(* PLC project PR_ModeManageNoMode_PLC, SiemensToBackhoff Siemens TIA Portal to Beckhoff TwinCAT PLCopen Converter 1.0 *)
(* stored: creationDateTime 2026-09-28T08:41:48.575973Z, modificationDateTime 2026-09-28T08:41:48.575973Z *)

FUNCTION_BLOCK PR_ModeManageNoMode

(* LD diagram, written out as Structured Text *)
(* Cycle Start delay validation
Cycle Start delay validation *)
inst_LT_11(pre := TRUE, in1 := TRUE, in2 := TRUE);
inst_GT_12(pre := TRUE, in1 := TRUE, in2 := TRUE);
inst_MOVE_13(in := TRUE, out1 => sCycleStartDelay);
inst_MOVE_14(in := TRUE, out1 => sCycleStartDelay);
(* Power ON reset Bit during initial power ON
Reset Active *)
sPowerOnReset := NOT iControlOn AND iFirstscan;
(* Control On pulse
#sControlOnPulse *)
inst_R_TRIG_20(in := TRUE, bit := TRUE);
sControlOnPulse := inst_R_TRIG_20.out;
(* Manual mode active
Man Mode *)
sManModeActive := iManMode AND sManModeActive AND NOT iAutoMode AND NOT sAutoRunningActive AND NOT sHomeRunningActive AND iManModeEnable AND NOT sPowerOnReset;
(* Waiting for cycle to start
Auto Mode *)
sWaitForCStart := iAutoMode AND NOT iManMode AND sWaitForCStart AND NOT iImmediateStop AND NOT sManModeActive AND NOT sAutoRunningActive AND iAutoModeEnable AND NOT sPowerOnReset;
(* CycleStartDelayTimer
CycleStartDelayTimer *)
CycleStartOnDelayTimer(IN := TRUE, PT := TRUE, ET := TRUE);
(* Drain,Dry,Cycle Stop Active
Drain,Dry,Cycle Stop Active *)
sDrainActive := true AND iDrainCycle AND true AND sDrainActive AND sAutoRunningActive AND NOT sPowerOnReset AND NOT iDryCycle AND NOT sDryCycleActive;
sDryCycleActive := true AND iDryCycle AND sWaitForCStart AND true AND sDryCycleActive AND NOT sManModeActive AND iAutoModeEnable AND NOT sPowerOnReset AND NOT iDrainCycle AND NOT sDrainActive;
sCycleStopActive := true AND iCycleStop AND true AND sAutoRunningActive AND iManMode AND true AND sCycleStopActive AND sAutoRunningActive AND NOT sPowerOnReset;
(* Auto running active
Auto Running *)
inst_UNKNOWN_75(IN := TRUE);
inst_UNKNOWN_77(IN := inst_UNKNOWN_75.Q AND NOT iDrainCompleted);
sAutoRunningActive := inst_UNKNOWN_77.Q AND NOT sDrainActive AND iAutoModeEnable AND NOT sPowerOnReset;
(* Home running active
Home Running Active *)
sHomeRunningActive := iHomePB AND qManModeActive AND sHomeRunningActive AND NOT iAutoMode AND NOT iHomeCompleted AND NOT sPowerOnReset AND iManModeEnable AND NOT iImmediateStop;
(* Resetting module to initial state
Module Reset *)
sModuleReset := NOT sManModeActive AND NOT sAutoRunningActive AND NOT sHomeRunningActive AND sManModeActive;
inst_R_TRIG_98(in := TRUE, bit := TRUE);
(* Message if machine is started without home conditions OK
Machine Not At Home if C Start Press *)
sMsgCStartandNoHome := iCycleStart AND sWaitForCStart AND NOT iHomeCompleted AND NOT iBypassHomeOption;
(* Message if manual mode selected during auto running
MsgManModeinAutoRunning *)
sMsgManModeinAutoRunning := sAutoRunningActive AND iManMode;
(* Outputs
Outputs *)
qManModeActive := sManModeActive;
qWaitForCStart := sWaitForCStart;
qDrainActive := sDrainActive;
qDryCycleActive := sDryCycleActive;
qCycleStopActive := sCycleStopActive;
qAutoRunningActive := sAutoRunningActive;
qHomeRunningActive := sHomeRunningActive;
qModuleReset := sModuleReset;
qMsgManModeinAutoRunning := sMsgManModeinAutoRunning;
qMsgCStartandNoHome := sMsgCStartandNoHome;
END_FUNCTION_BLOCK
